Fanuc KAREL source: KT00770.KL

PROGRAM KT00770
%NOLOCKGROUP
VAR
  S1: STRING[80]
  S2: STRING[80]
  OUT: INTEGER
BEGIN
  S1 = 'A'
  S2 = 'B'
  S1 = 'A'
  S2 = 'B'
  OUT = ACOS(S1)
END KT00770
